Yaskawa INFORM job: MAIN_1.JBI

/JOB
//NAME MAIN_1
//POS
///NPOS 80,0,0,0,0,0
///TOOL 9
///POSTYPE PULSE
///PULSE
C00000=0,0,0,0,0,0
C00001=0,3,-15,0,12,0
C00002=0,9,-17,0,-14,0
C00003=-29,47,0,27,25,-52
C00004=-29,56,0,39,18,-65
C00005=-29,47,0,27,25,-52
C00006=-13,39,14,20,15,-31
C00007=-13,51,14,59,6,-70
C00008=-13,39,14,20,15,-31
C00009=52,46,7,67,20,-93
C00010=52,46,7,67,20,-93
C00011=39,53,-5,56,30,-93
C00012=25,41,30,88,29,-142
C00013=25,41,30,88,29,-142
C00014=39,53,-5,56,30,-93
C00015=52,46,7,67,20,-93
C00016=52,46,7,67,20,-93
C00017=0,0,0,0,0,0
C00018=89,30,-6,-2,49,5
C00019=89,38,8,-3,27,6
C00020=70,42,-1,8,32,-22
C00021=69,41,1,0,42,-16
C00022=89,37,10,-3,39,6
C00023=88,25,24,-5,13,8
C00024=65,29,18,48,16,-63
C00025=64,15,13,24,32,-38
C00026=0,0,0,0,0,0
C00027=-68,24,27,38,36,-99
C00028=-68,31,28,47,30,-109
C00029=-69,36,24,48,30,-112
C00030=-70,38,21,46,31,-110
C00031=-71,40,17,44,33,-109
C00032=-73,42,14,42,34,-108
C00033=-74,43,11,40,36,-107
C00034=-76,44,8,39,38,-107
C00035=-77,46,6,37,39,-107
C00036=-79,47,4,36,40,-107
C00037=-81,47,3,35,42,-108
C00038=-83,48,2,35,43,-109
C00039=-85,48,1,34,43,-110
C00040=-87,48,1,34,44,-112
C00041=-88,48,2,33,45,-113
C00042=-90,47,3,33,45,-115
C00043=-92,46,4,33,45,-117
C00044=-94,45,6,33,45,-119
C00045=-95,44,9,33,44,-121
C00046=-97,43,11,34,44,-123
C00047=-98,41,14,34,43,-125
C00048=-100,40,17,34,42,-127
C00049=-101,38,21,35,41,-130
C00050=-102,36,24,36,40,-132
C00051=-102,34,28,37,38,-134
C00052=-102,34,28,37,39,-134
C00053=-103,33,32,38,37,-136
C00054=-103,31,35,40,36,-137
C00055=-102,29,39,41,35,-139
C00056=-101,27,42,43,33,-141
C00057=-100,26,45,46,32,-142
C00058=-98,24,48,48,31,-143
C00059=-96,23,50,51,29,-144
C00060=-93,22,52,54,28,-144
C00061=-90,21,53,57,27,-144
C00062=-87,21,54,60,27,-144
C00063=-84,21,54,62,26,-143
C00064=-80,21,53,64,25,-141
C00065=-77,22,52,65,25,-139
C00066=-75,23,50,66,25,-137
C00067=-72,24,48,65,24,-134
C00068=-71,26,45,64,25,-130
C00069=-69,27,42,61,25,-127
C00070=-69,29,38,59,25,-123
C00071=-68,31,35,56,26,-120
C00072=-68,33,31,53,27,-117
C00073=-69,35,28,51,28,-114
C00074=-69,36,24,48,30,-112
C00075=-70,36,18,41,34,-104
C00076=-70,30,17,35,40,-97
C00077=-29,47,0,27,25,-52
C00078=-29,56,0,39,18,-65
C00079=-29,47,0,27,25,-52
//INST
///DATE 2023/01/01 00:00
///COMM Generated using RoboDK
///ATTR SC,RW
///GROUP1 RB1
NOP
'Program generated by RoboDK v
'5.6.9 for RoboDK Industrial o
'n 26/02/2024 09:58:20
'Using nominal kinematics.
MOVJ C00000 VJ=50.00
MOVJ C00001 VJ=50.00
MOVL C00002 V=100.0
DOUT OT#(5) ON
DOUT OT#(5) ON
DOUT OT#(5) 0.5
DOUT OT#(5) true
DOUT OT#(5) ON
DOUT OT#(5) ON
DOUT OT#(5) 0.5
DOUT OT#(5) true
DOUT var val
DOUT var val
WAIT IN#(5)=ON
WAIT IN#(5)=ON
WAIT IN#(5)=0.5
WAIT IN#(5)=true
WAIT IN#(5)=ON T=0.10
WAIT var=val
WAIT var=val T=0.10
MSG "Message"
CALL JOB:REMOTE_
CODE_INSERT_172
'Insert Comment
'Using Frame Pick and Place (t
'argets wrt base):
'719.0,-664.0,0.0,0.0,0.0,0.0
'Tool 1 (Tool 1) should be clo
'se to:
'129.1,0.0,85.5,0.0,22.8,0.0
MOVJ C00003 VJ=100.0 ACC=100 DEC=100
MOVL C00004 V=100.0 ACC=100 DEC=100
DOUT OT#(5) ON
CALL JOB:PICK_PA
MOVL C00005 V=300.0 ACC=100 DEC=100
MOVL C00006 V=300.0 ACC=100 DEC=100
'MoveSearch command not implem
'ented
MOVL C00007 V=100.0 ACC=100 DEC=100
DOUT OT#(5) OFF
CALL JOB:PLACE_P
MOVL C00008 V=100.0 ACC=100 DEC=100
'Using Frame Circular (targets
' wrt base):
'577.7,392.2,0.0,0.0,0.0,39.0
MOVJ C00009 VJ=100.0 ACC=100 DEC=100
MOVC C00010 V=100.0 ACC=100 DEC=100 PL=8
MOVC C00011 V=100.0 ACC=100 DEC=100 PL=8
MOVC C00012 V=100.0 ACC=100 DEC=100 PL=8
MOVC C00013 V=100.0 ACC=100 DEC=100 PL=8
MOVC C00014 V=100.0 ACC=100 DEC=100 PL=8
MOVC C00015 V=100.0 ACC=100 DEC=100 PL=8
MOVL C00016 V=100.0 ACC=100 DEC=100
MOVJ C00017 VJ=100.0 ACC=100 DEC=100
'Using Frame Inspection (targe
'ts wrt base):
'0.0,782.7,377.6,0.0,0.0,0.0
MOVJ C00018 VJ=100.0 ACC=100 DEC=100
MOVL C00019 V=100.0 ACC=100 DEC=100
MOVL C00020 V=100.0 ACC=100 DEC=100
MOVL C00021 V=100.0 ACC=100 DEC=100
MOVL C00022 V=100.0 ACC=100 DEC=100
MOVL C00023 V=100.0 ACC=100 DEC=100
MOVL C00024 V=100.0 ACC=100 DEC=100
MOVL C00025 V=100.0 ACC=100 DEC=100
MOVJ C00026 VJ=100.0 ACC=100 DEC=100
CALL JOB:EVENT_P
'Using Frame Inspection (targe
'ts wrt base):
'13.6,-840.1,0.0,0.0,0.0,-90.0
'Show Tool 1
MOVJ C00027 VJ=100.0 ACC=100 DEC=100
CALL JOB:EVENT_P
MOVL C00028 V=1000.0 ACC=100 DEC=100
MOVL C00029 V=1000.0 ACC=100 DEC=100
CALL JOB:EVENT_P
MOVL C00030 V=50.0 ACC=100 DEC=100
MOVL C00031 V=50.0 ACC=100 DEC=100
MOVL C00032 V=50.0 ACC=100 DEC=100
MOVL C00033 V=50.0 ACC=100 DEC=100
MOVL C00034 V=50.0 ACC=100 DEC=100
MOVL C00035 V=50.0 ACC=100 DEC=100
MOVL C00036 V=50.0 ACC=100 DEC=100
MOVL C00037 V=50.0 ACC=100 DEC=100
MOVL C00038 V=50.0 ACC=100 DEC=100
MOVL C00039 V=50.0 ACC=100 DEC=100
MOVL C00040 V=50.0 ACC=100 DEC=100
MOVL C00041 V=50.0 ACC=100 DEC=100
MOVL C00042 V=50.0 ACC=100 DEC=100
MOVL C00043 V=50.0 ACC=100 DEC=100
MOVL C00044 V=50.0 ACC=100 DEC=100
MOVL C00045 V=50.0 ACC=100 DEC=100
MOVL C00046 V=50.0 ACC=100 DEC=100
MOVL C00047 V=50.0 ACC=100 DEC=100
MOVL C00048 V=50.0 ACC=100 DEC=100
MOVL C00049 V=50.0 ACC=100 DEC=100
MOVL C00050 V=50.0 ACC=100 DEC=100
MOVL C00051 V=50.0 ACC=100 DEC=100
MOVL C00052 V=50.0 ACC=100 DEC=100
MOVL C00053 V=50.0 ACC=100 DEC=100
MOVL C00054 V=50.0 ACC=100 DEC=100
MOVL C00055 V=50.0 ACC=100 DEC=100
MOVL C00056 V=50.0 ACC=100 DEC=100
MOVL C00057 V=50.0 ACC=100 DEC=100
MOVL C00058 V=50.0 ACC=100 DEC=100
MOVL C00059 V=50.0 ACC=100 DEC=100
MOVL C00060 V=50.0 ACC=100 DEC=100
MOVL C00061 V=50.0 ACC=100 DEC=100
MOVL C00062 V=50.0 ACC=100 DEC=100
MOVL C00063 V=50.0 ACC=100 DEC=100
MOVL C00064 V=50.0 ACC=100 DEC=100
MOVL C00065 V=50.0 ACC=100 DEC=100
MOVL C00066 V=50.0 ACC=100 DEC=100
MOVL C00067 V=50.0 ACC=100 DEC=100
MOVL C00068 V=50.0 ACC=100 DEC=100
MOVL C00069 V=50.0 ACC=100 DEC=100
MOVL C00070 V=50.0 ACC=100 DEC=100
MOVL C00071 V=50.0 ACC=100 DEC=100
MOVL C00072 V=50.0 ACC=100 DEC=100
MOVL C00073 V=50.0 ACC=100 DEC=100
MOVL C00074 V=50.0 ACC=100 DEC=100
CALL JOB:EVENT_P
MOVL C00075 V=1000.0 ACC=100 DEC=100
MOVL C00076 V=1000.0 ACC=100 DEC=100
CALL JOB:EVENT_P
CALL JOB:EVENT_P
'Using Frame Pick and Place (t
'argets wrt base):
'719.0,-664.0,0.0,0.0,0.0,0.0
MOVJ C00077 VJ=100.0 ACC=100 DEC=100
TIMER T=1.25
MOVL C00078 V=1000.0 ACC=100 DEC=100
WAIT IN#(1)=ON
MOVL C00079 V=1000.0 ACC=100 DEC=100
CALL JOB:PROG1_W
END
